(*
See the `Beckhoff Online Information System`__ or the `Beckhoff home page`__.

.. __: http://infosys.beckhoff.de/

.. __: http://beckhoff.de/
*)

FUNCTION_BLOCK FB_Libdoc_AnonymousHyperlinks
VAR_INPUT
    nVarA : INT;
    nVarB : INT;
END_VAR
VAR_OUTPUT
    nSum : INT;
END_VAR
VAR
END_VAR

END_FUNCTION_BLOCK

(* stored: Version 1.1.0.1, ProductVersion 3.1.4022.17
   POU FB_Libdoc_AnonymousHyperlinks: Id {1a8356c1-6a33-4dcd-a483-ad23079c7c24}, SpecialFunc None *)
